Fanuc KAREL source: KT00749.KL

PROGRAM KT00749
%NOLOCKGROUP
VAR
  I1: INTEGER
  I2: INTEGER
  OUT: REAL
BEGIN
  I1 = 2
  I2 = 3
  I1 = 2
  I2 = 3
  OUT = ABS(I1)
END KT00749
